(* IEC 61131-3 sources: trust-platform/examples/vat_pasteurizer/src, 8 files *)

(* ---- types.st ---- *)
(* The vat pasteurizer's types: its batch states, its recipe, its alarms, the signals of its plant,
   the operator's commands and what it shows the operator. *)

TYPE VatState :
(
    Idle := 0,
    Filling := 1,
    Heating := 2,
    Holding := 3,
    Cooling := 4,
    Draining := 5,
    Done := 6,
    Stopped := 7,
    Aborted := 8
);
END_TYPE

(* One product's heat treatment: the vat is filled to FillLevel, heated to PasteurTemp, held there
   for HoldTime and cooled to CoolTemp. *)
TYPE Recipe :
STRUCT
    Name : STRING[16];
    FillLevel : REAL;
    PasteurTemp : REAL;
    HoldTime : TIME;
    CoolTemp : REAL;
END_STRUCT
END_TYPE

(* One alarm: its condition now, raised and not yet reset, acknowledged by the operator. *)
TYPE AlarmEntry :
STRUCT
    Active : BOOL;
    Latched : BOOL;
    Acknowledged : BOOL;
END_STRUCT
END_TYPE

(* The plant's signals as the I/O wiring gives them: transmitters in raw counts, where 0 is 4 mA and
   27648 is 20 mA, switches and contactor feedbacks, and the outputs to valves, motors, the heater
   and the horn. A real installation binds these to its I/O; the bench's simulation drives them. *)
TYPE FieldSignals :
STRUCT
    LevelRaw : INT;
    TempRaw : INT;
    LevelHighHigh : BOOL;
    EmergencyStopOk : BOOL;
    InletOpen : BOOL;
    OutletOpen : BOOL;
    CoolingOpen : BOOL;
    AgitatorRunning : BOOL;
    PumpRunning : BOOL;
    InletValve : BOOL;
    OutletValve : BOOL;
    CoolingValve : BOOL;
    Agitator : BOOL;
    Pump : BOOL;
    HeaterPower : INT;
    Horn : BOOL;
END_STRUCT
END_TYPE

(* The operator's commands from the panel: each acts on its rising edge. *)
TYPE OperatorCommands :
STRUCT
    Start : BOOL;
    Stop : BOOL;
    Abort : BOOL;
    Reset : BOOL;
    Acknowledge : BOOL;
    RecipeIndex : INT := 1;
END_STRUCT
END_TYPE

(* What the panel shows: the batch's state and values, and the texts the panel's slow task builds. *)
TYPE VatStatus :
STRUCT
    State : VatState;
    Recipe : STRING[16];
    Level : REAL;
    Temperature : REAL;
    Setpoint : REAL;
    HeaterPower : REAL;
    HoldRemaining : TIME;
    StepTime : TIME;
    Batches : UDINT;
    ActiveAlarms : INT;
    Unacknowledged : INT;
    FirstOut : INT;
    StateText : STRING[48];
    AlarmText : STRING[40];
    BatchReport : STRING[64];
END_STRUCT
END_TYPE

(* ---- alarms.st ---- *)
(* The vat's alarms in the manner of ISA-18.2: an alarm is raised while its condition is present,
   stays latched until the operator has acknowledged it and its condition has cleared, and the first
   alarm raised since all were clear is kept as the first-out. The horn sounds while an alarm is
   unacknowledged. A critical alarm aborts the batch. *)

FUNCTION_BLOCK AlarmList
VAR_INPUT
    Conditions : ARRAY[1..12] OF BOOL;
    Acknowledge : BOOL;
END_VAR
VAR_OUTPUT
    Active : INT;
    Unacknowledged : INT;
    CriticalActive : BOOL;
    FirstOut : INT;
    Horn : BOOL;
    Raised : ARRAY[1..12] OF BOOL;
END_VAR
VAR
    Entries : ARRAY[1..12] OF AlarmEntry;
    AckEdge : R_TRIG;
    Index : INT;
    (* Emergency stop, level high-high, the two transmitters, over-temperature, agitator, inlet
       and outlet valve abort the batch; cooling valve, pump, heating timeout and a restarted hold
       warn. A variable, since the compiler cannot yet index a constant array by a variable. *)
    Critical : ARRAY[1..12] OF BOOL := [8(TRUE), 4(FALSE)];
END_VAR

AckEdge(CLK := Acknowledge);
Active := 0;
Unacknowledged := 0;
CriticalActive := FALSE;
FOR Index := 1 TO 12 DO
    IF Conditions[Index] AND NOT Entries[Index].Active THEN
        (* A new occurrence needs a new acknowledgement. *)
        Entries[Index].Latched := TRUE;
        Entries[Index].Acknowledged := FALSE;
        IF FirstOut = 0 THEN
            FirstOut := Index;
        END_IF;
    END_IF;
    Entries[Index].Active := Conditions[Index];
    IF AckEdge.Q THEN
        Entries[Index].Acknowledged := TRUE;
    END_IF;
    IF Entries[Index].Latched AND Entries[Index].Acknowledged AND NOT Entries[Index].Active THEN
        Entries[Index].Latched := FALSE;
    END_IF;
    Raised[Index] := Entries[Index].Latched;
    IF Entries[Index].Latched THEN
        Active := Active + 1;
        IF NOT Entries[Index].Acknowledged THEN
            Unacknowledged := Unacknowledged + 1;
        END_IF;
        IF Critical[Index] THEN
            CriticalActive := TRUE;
        END_IF;
    END_IF;
END_FOR;
IF Active = 0 THEN
    FirstOut := 0;
END_IF;
Horn := Unacknowledged > 0;
END_FUNCTION_BLOCK

(* ---- control.st ---- *)
NAMESPACE Control
TYPE PIDMode :
(
    Auto := 0,
    Manual := 1,
    Track := 2
);
END_TYPE

TYPE PIDAntiWindup :
(
    BackCalculation := 0,
    Combined := 1
);
END_TYPE

TYPE FilterOrder :
(
    FirstOrder := 0,
    SecondOrder := 1
);
END_TYPE

TYPE PIDParameters :
STRUCT
    ProportionalGain : LREAL;
    IntegralGain : LREAL;
    DerivativeGain : LREAL;
    ProportionalSetpointWeight : LREAL;
    DerivativeSetpointWeight : LREAL;
    Bias : LREAL;
    OutputMinimum : LREAL;
    OutputMaximum : LREAL;
    RateMinimum : LREAL;
    RateMaximum : LREAL;
    TrackingTime : LREAL;
    AntiWindup : PIDAntiWindup;
END_STRUCT
END_TYPE

TYPE PIDInitialState :
STRUCT
    Setpoint : LREAL;
    SetpointRate : LREAL;
    ProcessValue : LREAL;
    ProcessValueRate : LREAL;
    FeedForward : LREAL;
    NominalOutput : LREAL;
    SaturatedOutput : LREAL;
END_STRUCT
END_TYPE

TYPE PIDInput :
STRUCT
    Setpoint : LREAL;
    ProcessValue : LREAL;
    FeedForward : LREAL;
    ManualOutput : LREAL;
    TrackingOutput : LREAL;
    Mode : PIDMode;
    CycleTime : LREAL;
END_STRUCT
END_TYPE

TYPE LowPassParameters :
STRUCT
    TimeConstant : LREAL;
    Order : FilterOrder;
END_STRUCT
END_TYPE

FUNCTION_BLOCK PID
VAR
    ParametersValue : PIDParameters;
    StateValue : PIDInitialState;
END_VAR
(* truST simulation extension (specification 46, section 13.2): the measurement a simulated
   plant holds for this controller through a pid: feedback target, written between scans. A
   restart or a newly loaded program removes it. *)
VAR NON_RETAIN
    HeldMeasurement : LREAL;
    MeasurementHeld : BOOL;
END_VAR
(* truST observation extension (specification 45, section 3.1), beside GetState: the mode the
   last Update ran in, and whether Update has run since the start. A tool reads them; a restart
   clears them. *)
VAR NON_RETAIN
    ModeValue : PIDMode;
    ModeObserved : BOOL;
END_VAR

METHOD PUBLIC Configure
VAR_INPUT
    Parameters : PIDParameters;
END_VAR
ParametersValue := Parameters;
END_METHOD

METHOD PUBLIC Initialize
VAR_INPUT
    State : PIDInitialState;
END_VAR
StateValue := State;
END_METHOD

(* truST observation extension: a value copy, without a controller update. *)
METHOD PUBLIC GetState : PIDInitialState
GetState := StateValue;
END_METHOD

METHOD PUBLIC Update : LREAL
VAR_INPUT
    Input : PIDInput;
END_VAR
VAR
    Applied : PIDInput;
    LowerLimit : LREAL;
    UpperLimit : LREAL;
    SetpointRate : LREAL;
    ProcessValueRate : LREAL;
    NominalOutput : LREAL;
    SaturatedCandidate : LREAL;
    ProportionalIncrement : LREAL;
    IntegralIncrement : LREAL;
    DerivativeIncrement : LREAL;
    FeedForwardIncrement : LREAL;
    SaturationError : LREAL;
    ConditionalCorrection : LREAL;
    Output : LREAL;
END_VAR

(* The input the controller works on: Input, with the measurement a simulated plant holds as
   ProcessValue while one is held (simulation extension). *)
Applied := Input;
IF MeasurementHeld THEN
    Applied.ProcessValue := HeldMeasurement;
END_IF;

(* Rate limits are anchored to the actuator-facing saturated history. *)
LowerLimit := MAX(
    ParametersValue.OutputMinimum,
    StateValue.SaturatedOutput + Applied.CycleTime * ParametersValue.RateMinimum
);
UpperLimit := MIN(
    ParametersValue.OutputMaximum,
    StateValue.SaturatedOutput + Applied.CycleTime * ParametersValue.RateMaximum
);

SetpointRate := (Applied.Setpoint - StateValue.Setpoint) / Applied.CycleTime;
ProcessValueRate := (Applied.ProcessValue - StateValue.ProcessValue) / Applied.CycleTime;

IF Applied.Mode = Track THEN
    StateValue.NominalOutput := Applied.TrackingOutput;
END_IF;

IF Applied.Mode = Manual THEN
    NominalOutput := Applied.ManualOutput;
ELSE
    IF ParametersValue.IntegralGain = LREAL#0.0 THEN
        NominalOutput := ParametersValue.Bias
            + ParametersValue.ProportionalGain * (Applied.Setpoint - Applied.ProcessValue)
            + ParametersValue.DerivativeGain
                * (ParametersValue.DerivativeSetpointWeight * SetpointRate - ProcessValueRate)
            + Applied.FeedForward;
    ELSE
        ProportionalIncrement := ParametersValue.ProportionalGain
            * (ParametersValue.ProportionalSetpointWeight
                * (Applied.Setpoint - StateValue.Setpoint)
                - (Applied.ProcessValue - StateValue.ProcessValue));
        IntegralIncrement := ParametersValue.IntegralGain * Applied.CycleTime
            * (Applied.Setpoint - Applied.ProcessValue);
        DerivativeIncrement := ParametersValue.DerivativeGain
            * (ParametersValue.DerivativeSetpointWeight
                * (SetpointRate - StateValue.SetpointRate)
                - (ProcessValueRate - StateValue.ProcessValueRate));
        FeedForwardIncrement := Applied.FeedForward - StateValue.FeedForward;

        NominalOutput := StateValue.NominalOutput
            + ProportionalIncrement
            + IntegralIncrement
            + DerivativeIncrement
            + FeedForwardIncrement;
        SaturatedCandidate := MAX(MIN(NominalOutput, UpperLimit), LowerLimit);
        IF ParametersValue.AntiWindup = Combined THEN
            SaturationError := NominalOutput - SaturatedCandidate;
            IF IntegralIncrement * SaturationError > LREAL#0.0 THEN
                ConditionalCorrection := MIN(ABS(IntegralIncrement), ABS(SaturationError));
                IF SaturationError > LREAL#0.0 THEN
                    NominalOutput := NominalOutput - ConditionalCorrection;
                ELSE
                    NominalOutput := NominalOutput + ConditionalCorrection;
                END_IF;
            END_IF;
            (* Listing 5 deliberately reuses the candidate from before the correction. *)
            NominalOutput := NominalOutput
                - MIN(Applied.CycleTime / ParametersValue.TrackingTime, LREAL#1.0)
                    * (NominalOutput - SaturatedCandidate);
        ELSE
            NominalOutput := NominalOutput
                - Applied.CycleTime / ParametersValue.TrackingTime
                    * (NominalOutput - SaturatedCandidate);
        END_IF;
    END_IF;
END_IF;

StateValue.NominalOutput := NominalOutput;
Output := MAX(MIN(NominalOutput, UpperLimit), LowerLimit);
StateValue.SaturatedOutput := Output;
StateValue.Setpoint := Applied.Setpoint;
StateValue.SetpointRate := SetpointRate;
StateValue.ProcessValue := Applied.ProcessValue;
StateValue.ProcessValueRate := ProcessValueRate;
StateValue.FeedForward := Applied.FeedForward;
(* Observation extension: the mode this call ran in. *)
ModeValue := Applied.Mode;
ModeObserved := TRUE;
Update := Output;
END_METHOD
END_FUNCTION_BLOCK

FUNCTION_BLOCK LowPass
VAR
    ParametersValue : LowPassParameters;
    Stage1 : LREAL;
    Stage2 : LREAL;
END_VAR

METHOD PUBLIC Configure
VAR_INPUT
    Parameters : LowPassParameters;
END_VAR
ParametersValue := Parameters;
END_METHOD

METHOD PUBLIC Initialize
VAR_INPUT
    Input : LREAL;
END_VAR
Stage1 := Input;
Stage2 := Input;
END_METHOD

METHOD PUBLIC Update : LREAL
VAR_INPUT
    Input : LREAL;
    CycleTime : LREAL;
END_VAR
VAR
    Coefficient : LREAL;
    NextStage1 : LREAL;
    NextStage2 : LREAL;
END_VAR

Coefficient := CycleTime / (ParametersValue.TimeConstant + LREAL#0.5 * CycleTime);
NextStage1 := Stage1 + Coefficient * (Input - Stage1);
Stage1 := NextStage1;

IF ParametersValue.Order = SecondOrder THEN
    NextStage2 := Stage2 + Coefficient * (NextStage1 - Stage2);
    Stage2 := NextStage2;
    Update := NextStage2;
ELSE
    Update := NextStage1;
END_IF;
END_METHOD
END_FUNCTION_BLOCK
END_NAMESPACE

(* ---- equipment.st ---- *)
(* The vat's equipment: a valve or a motor with its feedback, and a 4-20 mA transmitter. *)

(* A valve with an open limit switch, or a motor with its contactor's running feedback: it is
   driven while it is commanded and its interlock allows it. A feedback that does not follow the
   output within the supervision time is a fault, which keeps it off until it is reset. *)
FUNCTION_BLOCK Actuator
VAR_INPUT
    Command : BOOL;
    Interlock : BOOL := TRUE;
    Feedback : BOOL;
    Reset : BOOL;
    SupervisionTime : TIME := T#3s;
END_VAR
VAR_OUTPUT
    Output : BOOL;
    Fault : BOOL;
END_VAR
VAR
    Mismatch : TON;
END_VAR

IF Reset THEN
    Fault := FALSE;
END_IF;
Output := Command AND Interlock AND NOT Fault;
Mismatch(IN := Output <> Feedback, PT := SupervisionTime);
IF Mismatch.Q THEN
    Fault := TRUE;
    Output := FALSE;
END_IF;
END_FUNCTION_BLOCK

(* A 4-20 mA transmitter read as raw counts, 0 at 4 mA and 27648 at 20 mA, scaled to its range.
   Below 3.6 mA or above 21 mA the loop is broken or shorted (NAMUR NE 43): the value is then a fault
   and keeps its last good reading. *)
FUNCTION_BLOCK AnalogInput
VAR_INPUT
    Raw : INT;
    RangeLow : REAL;
    RangeHigh : REAL;
END_VAR
VAR_OUTPUT
    Value : REAL;
    Fault : BOOL;
END_VAR

Fault := Raw < -691 OR Raw > 29376;
IF NOT Fault THEN
    Value := RangeLow + (RangeHigh - RangeLow) * INT_TO_REAL(Raw) / 27648.0;
END_IF;
END_FUNCTION_BLOCK

(* ---- config.st ---- *)
(* The vat pasteurizer on one controller: the batch control every 10 ms, the simulated plant every
   20 ms and the panel's texts every 500 ms. The lamps are the bench's outputs; the register map is
   what a panel or a SCADA system reads over the network. *)
CONFIGURATION VatPasteurizer
VAR_GLOBAL
    Io : FieldSignals;
    Panel : OperatorCommands;
    Status : VatStatus;
END_VAR
RESOURCE Plc ON PLC
    TASK ControlTask (INTERVAL := T#10ms, PRIORITY := 1);
    TASK SimulationTask (INTERVAL := T#20ms, PRIORITY := 2);
    TASK PanelTask (INTERVAL := T#500ms, PRIORITY := 3);
    PROGRAM Vat WITH ControlTask : VatControl;
    PROGRAM Plant WITH SimulationTask : PlantSimulation;
    PROGRAM Texts WITH PanelTask : PanelTexts;
END_RESOURCE
VAR_CONFIG
    Vat.LampRunning AT %QX0.0 : BOOL;
    Vat.LampWarning AT %QX0.1 : BOOL;
    Vat.LampAlarm AT %QX0.2 : BOOL;
    Vat.RegState AT %MW0 : INT;
    Vat.RegAlarms AT %MW2 : INT;
    Vat.RegTemperature AT %MD4 : DINT;
    Vat.RegLevel AT %MD8 : DINT;
    Vat.RegBatches AT %MD12 : UDINT;
END_VAR
END_CONFIGURATION

(* ---- panel.st ---- *)
(* The operator panel's texts, built in the slow panel task from the values the control task gives
   the panel: the state of the batch with its live values, the most important alarm, and a report
   line for the last batch. *)

(* The number of a state in the panel's register map. *)
FUNCTION StateCode : INT
VAR_INPUT
    State : VatState;
END_VAR
CASE State OF
    VatState#Idle: StateCode := 0;
    VatState#Filling: StateCode := 1;
    VatState#Heating: StateCode := 2;
    VatState#Holding: StateCode := 3;
    VatState#Cooling: StateCode := 4;
    VatState#Draining: StateCode := 5;
    VatState#Done: StateCode := 6;
    VatState#Stopped: StateCode := 7;
    VatState#Aborted: StateCode := 8;
END_CASE;
END_FUNCTION

(* A value with one decimal, as a panel shows it: 63.2. *)
FUNCTION OneDecimal : STRING[12]
VAR_INPUT
    Value : REAL;
END_VAR
VAR
    Tenths : DINT;
END_VAR
Tenths := REAL_TO_DINT(ABS(Value) * 10.0);
OneDecimal := CONCAT(DINT_TO_STRING(Tenths / 10), '.', DINT_TO_STRING(Tenths MOD 10));
IF Value < 0.0 THEN
    OneDecimal := CONCAT('-', OneDecimal);
END_IF;
END_FUNCTION

(* A duration as minutes and seconds: 17:05. *)
FUNCTION MinutesSeconds : STRING[12]
VAR_INPUT
    Duration : TIME;
END_VAR
VAR
    Seconds : UDINT;
END_VAR
Seconds := DWORD_TO_UDINT(TIME_TO_DWORD(Duration)) / 1000;
IF Seconds MOD 60 < 10 THEN
    MinutesSeconds := CONCAT(UDINT_TO_STRING(Seconds / 60), ':0', UDINT_TO_STRING(Seconds MOD 60));
ELSE
    MinutesSeconds := CONCAT(UDINT_TO_STRING(Seconds / 60), ':', UDINT_TO_STRING(Seconds MOD 60));
END_IF;
END_FUNCTION

PROGRAM PanelTexts
VAR_EXTERNAL
    Status : VatStatus;
END_VAR
VAR
    LastBatches : UDINT;
    (* In the order of the alarm conditions of VatControl. A variable, since the compiler cannot
       yet index a constant array by a variable. *)
    AlarmTexts : ARRAY[1..12] OF STRING[28] := [
        'Emergency stop',
        'Level high-high',
        'Level transmitter fault',
        'Temperature sensor fault',
        'Over-temperature',
        'Agitator fault',
        'Inlet valve fault',
        'Outlet valve fault',
        'Cooling valve fault',
        'Drain pump fault',
        'Heating takes too long',
        'Hold restarted: too cool'
    ];
END_VAR

CASE Status.State OF
    VatState#Idle:
        Status.StateText := CONCAT('Ready, recipe ', Status.Recipe);
    VatState#Filling:
        Status.StateText := CONCAT('Filling ', OneDecimal(Value := Status.Level), ' %');
    VatState#Heating:
        Status.StateText := CONCAT('Heating ', OneDecimal(Value := Status.Temperature), ' C to ',
            OneDecimal(Value := Status.Setpoint), ' C');
    VatState#Holding:
        Status.StateText := CONCAT('Holding ', OneDecimal(Value := Status.Temperature), ' C, ',
            MinutesSeconds(Duration := Status.HoldRemaining), ' left');
    VatState#Cooling:
        Status.StateText := CONCAT('Cooling ', OneDecimal(Value := Status.Temperature), ' C');
    VatState#Draining:
        Status.StateText := CONCAT('Draining ', OneDecimal(Value := Status.Level), ' %');
    VatState#Done:
        Status.StateText := 'Batch complete';
    VatState#Stopped:
        Status.StateText := CONCAT('Stopped for ', MinutesSeconds(Duration := Status.StepTime),
            ', Start resumes');
    VatState#Aborted:
        Status.StateText := 'Aborted: clear the alarms, then Reset';
END_CASE;

IF Status.FirstOut > 0 THEN
    Status.AlarmText := AlarmTexts[Status.FirstOut];
ELSE
    Status.AlarmText := '';
END_IF;

IF Status.Batches <> LastBatches THEN
    Status.BatchReport := CONCAT('Batch ', UDINT_TO_STRING(Status.Batches), ': ', Status.Recipe,
        ' pasteurized at ', OneDecimal(Value := Status.Setpoint), ' C');
    LastBatches := Status.Batches;
END_IF;
END_PROGRAM

(* ---- simulation.st ---- *)
(* The plant and its operator, simulated in a task of their own so that the vat runs whole batches
   on a bench with no plant wired. A real installation drops this program and wires FieldSignals to
   its I/O.

   The vat: the inlet fills it at 2 %/s with product at 8 C; the outlet with the drain pump running
   empties it at 2.5 %/s. The jacket heats the product at up to 0.25 C/s in a vat filled to 80 %,
   faster in a vat that holds less, and half as fast without agitation; the cooling water draws it
   towards 4 C with a time constant of 100 s; it loses heat towards 20 C slowly. Valves open
   1.5 s after they are commanded, motors run 0.5 s after they are started.

   The operator starts the bench recipe when the vat is idle, acknowledges a new alarm after 5 s and
   resets an aborted batch once its alarms are acknowledged. Every second batch the steam supply
   fails for 20 s while the vat holds, which restarts the hold; every third batch the agitator's
   contactor drops for 4 s while the vat heats, which aborts the batch. *)
PROGRAM PlantSimulation
VAR_EXTERNAL
    Io : FieldSignals;
    Panel : OperatorCommands;
    Status : VatStatus;
END_VAR
VAR
    LevelPercent : REAL := 0.0;
    Temp : REAL := 8.0;
    Seconds : REAL;
    Now : TIME;
    LastTime : TIME;
    Started : BOOL;
    InletTravel : TON;
    OutletTravel : TON;
    CoolingTravel : TON;
    AgitatorStart : TON;
    PumpStart : TON;
    HeatRate : REAL;
    (* The operator: a press lasts 0.3 s, as a finger on a button does. *)
    WaitIdle : TON;
    WaitAlarm : TON;
    WaitAborted : TON;
    Press : TP;
    Pressing : INT;
    (* The disturbances, by the batch they happen in and the time in the step. *)
    SimulatedBatches : UDINT;
    LastState : VatState := VatState#Idle;
    SteamFailure : BOOL;
    ContactorDrop : BOOL;
END_VAR

Now := TIME();
IF NOT Started THEN
    LastTime := Now;
    Started := TRUE;
END_IF;
Seconds := UDINT_TO_REAL(DWORD_TO_UDINT(TIME_TO_DWORD(Now - LastTime))) / 1000.0;
LastTime := Now;

(* The equipment follows its outputs. *)
InletTravel(IN := Io.InletValve, PT := T#1500ms);
OutletTravel(IN := Io.OutletValve, PT := T#1500ms);
CoolingTravel(IN := Io.CoolingValve, PT := T#1500ms);
AgitatorStart(IN := Io.Agitator, PT := T#500ms);
PumpStart(IN := Io.Pump, PT := T#500ms);
IF Status.State <> LastState THEN
    IF Status.State = VatState#Filling THEN
        SimulatedBatches := SimulatedBatches + 1;
    END_IF;
    LastState := Status.State;
END_IF;
SteamFailure := SimulatedBatches MOD 2 = 0 AND Status.State = VatState#Holding
    AND Status.StepTime >= T#10s AND Status.StepTime < T#30s;
ContactorDrop := SimulatedBatches MOD 3 = 0 AND Status.State = VatState#Heating
    AND Status.StepTime >= T#20s AND Status.StepTime < T#24s;
Io.InletOpen := InletTravel.Q;
Io.OutletOpen := OutletTravel.Q;
Io.CoolingOpen := CoolingTravel.Q;
Io.AgitatorRunning := AgitatorStart.Q AND NOT ContactorDrop;
Io.PumpRunning := PumpStart.Q;
Io.EmergencyStopOk := TRUE;

(* The vat's level and its product's temperature. *)
IF Io.InletOpen THEN
    LevelPercent := LevelPercent + 2.0 * Seconds;
    IF LevelPercent > 0.0 THEN
        Temp := Temp + (8.0 - Temp) * 2.0 * Seconds / LevelPercent;
    END_IF;
END_IF;
IF Io.OutletOpen AND Io.PumpRunning THEN
    LevelPercent := MAX(LevelPercent - 2.5 * Seconds, 0.0);
END_IF;
IF NOT SteamFailure AND LevelPercent > 5.0 THEN
    HeatRate := 0.25 * 80.0 / LevelPercent;
    IF NOT Io.AgitatorRunning THEN
        HeatRate := HeatRate * 0.5;
    END_IF;
    Temp := Temp + INT_TO_REAL(Io.HeaterPower) / 27648.0 * HeatRate * Seconds;
END_IF;
IF Io.CoolingOpen THEN
    Temp := Temp + (4.0 - Temp) * 0.01 * Seconds;
END_IF;
Temp := Temp + (20.0 - Temp) * 0.0005 * Seconds;
IF SteamFailure THEN
    (* The jacket's condensate cools the product. *)
    Temp := Temp - 0.08 * Seconds;
END_IF;
Io.LevelRaw := REAL_TO_INT(LevelPercent / 100.0 * 27648.0);
Io.TempRaw := REAL_TO_INT(Temp / 100.0 * 27648.0);
Io.LevelHighHigh := LevelPercent > 95.0;

(* The operator. *)
WaitIdle(IN := Status.State = VatState#Idle, PT := T#5s);
WaitAlarm(IN := Status.Unacknowledged > 0, PT := T#5s);
WaitAborted(IN := Status.State = VatState#Aborted AND Status.Unacknowledged = 0, PT := T#5s);
IF NOT Press.Q THEN
    IF Pressing > 0 THEN
        (* The press has ended: the finger leaves the button for one scan, so that the next press
           is a new rising edge. *)
        Pressing := 0;
    ELSIF WaitAlarm.Q THEN
        Pressing := 3;
    ELSIF WaitAborted.Q THEN
        Pressing := 2;
    ELSIF WaitIdle.Q THEN
        Pressing := 1;
    END_IF;
END_IF;
Press(IN := Pressing > 0, PT := T#300ms);
Panel.RecipeIndex := 2;
Panel.Start := Press.Q AND Pressing = 1;
Panel.Reset := Press.Q AND Pressing = 2;
Panel.Acknowledge := Press.Q AND Pressing = 3;
END_PROGRAM

(* ---- vat.st ---- *)
USING Control;

(* The vat pasteurizer's batch control, run in the control task. It reads the transmitters, runs the
   batch's state machine, the product temperature loop (Control.PID on the jacket heater), the
   valves and motors, raises the alarms and drives the outputs and the panel's values.

   A batch fills the vat to the recipe's level, heats the product with the agitator running, holds
   it at the pasteurizing temperature for the hold time, cools it and drains it. The hold counts
   only while the product stays within HoldBand of the pasteurizing temperature: if it falls below,
   the hold starts again, as the rules for a vat pasteurizer require. Stop pauses a batch and Start
   resumes it, a hold from its beginning. A critical alarm or Abort aborts the batch; Reset, once no
   critical alarm is left, drains a vat that holds product, else returns to Idle. *)
PROGRAM VatControl
VAR_EXTERNAL
    Io : FieldSignals;
    Panel : OperatorCommands;
    Status : VatStatus;
END_VAR
VAR
    State : VatState := VatState#Idle;
    PreviousState : VatState := VatState#Idle;
    Interrupted : VatState := VatState#Idle;
    Recipes : ARRAY[1..2] OF Recipe := [
        (Name := 'Milk LTLT', FillLevel := 80.0, PasteurTemp := 63.0, HoldTime := T#30m,
            CoolTemp := 6.0),
        (Name := 'Bench test', FillLevel := 40.0, PasteurTemp := 63.0, HoldTime := T#60s,
            CoolTemp := 30.0)
    ];
    Active : Recipe;
    Level : AnalogInput;
    Temperature : AnalogInput;
    TempFilter : Control.LowPass;
    FilterParameters : Control.LowPassParameters := (
        TimeConstant := LREAL#2.0,
        Order := FilterOrder#FirstOrder
    );
    Heater : Control.PID;
    HeaterParameters : Control.PIDParameters := (
        ProportionalGain := LREAL#8.0,
        IntegralGain := LREAL#0.08,
        DerivativeGain := LREAL#0.0,
        ProportionalSetpointWeight := LREAL#1.0,
        DerivativeSetpointWeight := LREAL#0.0,
        Bias := LREAL#0.0,
        OutputMinimum := LREAL#0.0,
        OutputMaximum := LREAL#100.0,
        RateMinimum := LREAL#-20.0,
        RateMaximum := LREAL#20.0,
        TrackingTime := LREAL#5.0,
        AntiWindup := PIDAntiWindup#Combined
    );
    HeaterInitial : Control.PIDInitialState;
    HeaterInput : Control.PIDInput;
    HeaterOutput : LREAL;
    Inlet : Actuator;
    Outlet : Actuator;
    Cooling : Actuator;
    Agitator : Actuator;
    Pump : Actuator;
    Alarms : AlarmList;
    Conditions : ARRAY[1..12] OF BOOL;
    StartEdge : R_TRIG;
    StopEdge : R_TRIG;
    AbortEdge : R_TRIG;
    ResetEdge : R_TRIG;
    ResetRequested : BOOL;
    StepTimer : TON;
    HoldTimer : TON;
    HeatingTimeout : TON;
    Initialized : BOOL;
    Now : TIME;
    LastTime : TIME;
    LoopElapsed : TIME;
    HoldRestarted : BOOL;
    InBatch : BOOL;
    (* The lamps of the panel, and the panel's register map. *)
    LampRunning : BOOL;
    LampWarning : BOOL;
    LampAlarm : BOOL;
    RegState : INT;
    RegTemperature : DINT;
    RegLevel : DINT;
    RegAlarms : INT;
    RegBatches : UDINT;
END_VAR
VAR RETAIN
    Batches : UDINT;
END_VAR
VAR CONSTANT
    (* The temperature loop's sample period. *)
    LoopPeriod : TIME := T#100ms;
    HoldBand : REAL := 0.5;
    OverTemperature : REAL := 75.0;
    (* Below this level the vat counts as empty. *)
    EmptyLevel : REAL := 2.0;
    (* Below this level the agitator's blades are not covered. *)
    AgitatorLevel : REAL := 20.0;
    MaxHeatingTime : TIME := T#15m;
    LoopAuto : Control.PIDMode := PIDMode#Auto;
    LoopManual : Control.PIDMode := PIDMode#Manual;
END_VAR

(* The transmitters. *)
Level(Raw := Io.LevelRaw, RangeLow := 0.0, RangeHigh := 100.0);
Temperature(Raw := Io.TempRaw, RangeLow := 0.0, RangeHigh := 100.0);
Now := TIME();
IF NOT Initialized THEN
    TempFilter.Configure(Parameters := FilterParameters);
    TempFilter.Initialize(Input := REAL_TO_LREAL(Temperature.Value));
    Heater.Configure(Parameters := HeaterParameters);
    HeaterInitial.Setpoint := REAL_TO_LREAL(Temperature.Value);
    HeaterInitial.ProcessValue := HeaterInitial.Setpoint;
    Heater.Initialize(State := HeaterInitial);
    Active := Recipes[1];
    LastTime := Now;
    Initialized := TRUE;
END_IF;

(* The operator's commands act on their rising edges. *)
StartEdge(CLK := Panel.Start);
StopEdge(CLK := Panel.Stop);
AbortEdge(CLK := Panel.Abort);
ResetEdge(CLK := Panel.Reset);

(* The alarms, in the order of AlarmList's critical table and of the panel's texts. *)
Conditions[1] := NOT Io.EmergencyStopOk;
Conditions[2] := Io.LevelHighHigh;
Conditions[3] := Level.Fault;
Conditions[4] := Temperature.Fault;
Conditions[5] := Temperature.Value > OverTemperature;
Conditions[6] := Agitator.Fault;
Conditions[7] := Inlet.Fault;
Conditions[8] := Outlet.Fault;
Conditions[9] := Cooling.Fault;
Conditions[10] := Pump.Fault;
Conditions[11] := HeatingTimeout.Q;
Conditions[12] := HoldRestarted;
Alarms(Conditions := Conditions, Acknowledge := Panel.Acknowledge);

(* The state machine. *)
CASE State OF
    VatState#Filling, VatState#Heating, VatState#Holding, VatState#Cooling, VatState#Draining:
        InBatch := TRUE;
ELSE
    InBatch := FALSE;
END_CASE;
IF (Alarms.CriticalActive OR AbortEdge.Q) AND InBatch THEN
    State := VatState#Aborted;
ELSIF StopEdge.Q AND InBatch THEN
    Interrupted := State;
    State := VatState#Stopped;
END_IF;

CASE State OF
    VatState#Idle:
        IF StartEdge.Q AND NOT Alarms.CriticalActive THEN
            Active := Recipes[LIMIT(1, Panel.RecipeIndex, 2)];
            State := VatState#Filling;
        END_IF;
    VatState#Filling:
        IF Level.Value >= Active.FillLevel THEN
            State := VatState#Heating;
        END_IF;
    VatState#Heating:
        (* The loop approaches its setpoint from below, so the hold starts within its band. *)
        IF Temperature.Value >= Active.PasteurTemp - HoldBand THEN
            State := VatState#Holding;
        END_IF;
    VatState#Holding:
        IF HoldTimer.Q THEN
            State := VatState#Cooling;
        END_IF;
    VatState#Cooling:
        IF Temperature.Value <= Active.CoolTemp THEN
            State := VatState#Draining;
        END_IF;
    VatState#Draining:
        (* The pump runs on for 5 s after the vat reads empty. *)
        IF Level.Value > EmptyLevel THEN
            StepTimer(IN := FALSE);
        ELSIF StepTimer.ET >= T#5s THEN
            State := VatState#Done;
        END_IF;
    VatState#Done:
        IF StepTimer.ET >= T#3s THEN
            State := VatState#Idle;
        END_IF;
    VatState#Stopped:
        IF StartEdge.Q AND NOT Alarms.CriticalActive THEN
            State := Interrupted;
        END_IF;
    VatState#Aborted:
        IF ResetEdge.Q THEN
            ResetRequested := TRUE;
        END_IF;
        IF ResetRequested AND NOT Alarms.CriticalActive THEN
            ResetRequested := FALSE;
            IF Level.Value > EmptyLevel THEN
                State := VatState#Draining;
            ELSE
                State := VatState#Idle;
            END_IF;
        END_IF;
END_CASE;

IF State <> PreviousState THEN
    StepTimer(IN := FALSE);
    IF State = VatState#Done THEN
        Batches := Batches + 1;
    END_IF;
    PreviousState := State;
END_IF;
StepTimer(IN := TRUE, PT := T#24h);

(* The hold counts only while the product is hot enough; a fall below restarts it. *)
HoldRestarted := State = VatState#Holding
    AND Temperature.Value < Active.PasteurTemp - HoldBand
    AND HoldTimer.ET > T#0s;
HoldTimer(IN := State = VatState#Holding AND Temperature.Value >= Active.PasteurTemp - HoldBand,
    PT := Active.HoldTime);
HeatingTimeout(IN := State = VatState#Heating, PT := MaxHeatingTime);

(* The valves and motors; the emergency stop drops them all. *)
Inlet(Command := State = VatState#Filling,
    Interlock := Io.EmergencyStopOk AND NOT Io.LevelHighHigh,
    Feedback := Io.InletOpen, Reset := ResetEdge.Q);
Agitator(Command := State = VatState#Heating OR State = VatState#Holding
        OR State = VatState#Cooling,
    Interlock := Io.EmergencyStopOk AND Level.Value > AgitatorLevel,
    Feedback := Io.AgitatorRunning, Reset := ResetEdge.Q, SupervisionTime := T#2s);
Cooling(Command := State = VatState#Cooling, Interlock := Io.EmergencyStopOk,
    Feedback := Io.CoolingOpen, Reset := ResetEdge.Q);
Outlet(Command := State = VatState#Draining, Interlock := Io.EmergencyStopOk,
    Feedback := Io.OutletOpen, Reset := ResetEdge.Q);
Pump(Command := State = VatState#Draining AND Io.OutletOpen,
    Interlock := Io.EmergencyStopOk, Feedback := Io.PumpRunning, Reset := ResetEdge.Q,
    SupervisionTime := T#2s);

(* The temperature loop runs at its own sample period, on the time that has actually passed. *)
LoopElapsed := LoopElapsed + (Now - LastTime);
LastTime := Now;
IF LoopElapsed >= LoopPeriod THEN
    HeaterInput.CycleTime := UDINT_TO_LREAL(DWORD_TO_UDINT(TIME_TO_DWORD(LoopElapsed))) / LREAL#1000.0;
    HeaterInput.ProcessValue := TempFilter.Update(
        Input := REAL_TO_LREAL(Temperature.Value),
        CycleTime := HeaterInput.CycleTime
    );
    HeaterInput.Setpoint := REAL_TO_LREAL(Active.PasteurTemp);
    IF State = VatState#Heating OR State = VatState#Holding THEN
        HeaterInput.Mode := LoopAuto;
    ELSE
        HeaterInput.Mode := LoopManual;
    END_IF;
    HeaterInput.ManualOutput := LREAL#0.0;
    HeaterOutput := Heater.Update(Input := HeaterInput);
    LoopElapsed := T#0s;
END_IF;

(* The outputs: heating without agitation would scorch the product. *)
Io.InletValve := Inlet.Output;
Io.OutletValve := Outlet.Output;
Io.CoolingValve := Cooling.Output;
Io.Agitator := Agitator.Output;
Io.Pump := Pump.Output;
IF Agitator.Output AND Io.AgitatorRunning THEN
    Io.HeaterPower := REAL_TO_INT(LREAL_TO_REAL(HeaterOutput) * 276.48);
ELSE
    Io.HeaterPower := 0;
END_IF;
Io.Horn := Alarms.Horn;
LampRunning := InBatch;
LampWarning := Alarms.Active > 0 AND NOT Alarms.CriticalActive;
LampAlarm := Alarms.CriticalActive;

(* The panel's values and register map. *)
Status.State := State;
Status.Recipe := Active.Name;
Status.Level := Level.Value;
Status.Temperature := Temperature.Value;
Status.Setpoint := Active.PasteurTemp;
Status.HeaterPower := LREAL_TO_REAL(HeaterOutput);
IF State = VatState#Holding THEN
    Status.HoldRemaining := Active.HoldTime - HoldTimer.ET;
ELSE
    Status.HoldRemaining := T#0s;
END_IF;
Status.StepTime := StepTimer.ET;
Status.Batches := Batches;
Status.ActiveAlarms := Alarms.Active;
Status.Unacknowledged := Alarms.Unacknowledged;
Status.FirstOut := Alarms.FirstOut;
RegState := StateCode(State := State);
RegTemperature := REAL_TO_DINT(Temperature.Value * 10.0);
RegLevel := REAL_TO_DINT(Level.Value * 10.0);
RegAlarms := Alarms.Active;
RegBatches := Batches;
END_PROGRAM
